FUNCTION SumFunction (* Adds two input values *)
  (* Standard: 61499-1; Description: Copyright (c) 2026 Martin Erich Jobst This program and the accompanying materials are made available under the terms of the Eclipse Public License 2.0 which is available at https://www.eclipse.org/legal/epl-2.0/ SPDX-License-Identifier: EPL-2.0 *)
  (* Version 1.0, 2026-10-23, Martin Jobst *)
  {SET_ATTRIBUTE(IntegerAttribute, 9)}
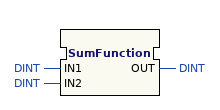
  VAR_INPUT
    IN1 : DINT;
    IN2 : DINT;
  END_VAR
  VAR_OUTPUT
    OUT : DINT;
  END_VAR
  BODY IN ST:
OUT := IN1 + IN2;
  END_BODY
END_FUNCTION
